(* Tests FB_Span.cloneTo, which processors use to keep a span that must outlive the original.
   A running span's context is taken through FB_Tracer.getSpanContext, tested in FB_TestTracer. *)
FUNCTION_BLOCK FB_TestSpan EXTENDS FB_TestSuite

THIS^.testCloneToCopiesEveryMember();
THIS^.testCloneToRejectsAssignedDestination();

(* cloneTo gives the copy its own copy of every member, so it outlives the source. *)
METHOD testCloneToCopiesEveryMember : REFERENCE TO FB_Test
VAR
	resource: FB_Resource('');
	idGenerator: FB_MockIdGenerator;
	provider: FB_TracerProvider_ForInspection(resource:=resource, idGenerator:=idGenerator, sampler:=TcOtlp_GVL.defaultSampler);
	scope: FB_InstrumentationScope('tracer.test', '1.0.0', '');
	tracer: FB_Tracer(scope:=scope, provider:=provider);
	pParent: POINTER TO FB_Span;
	pContext: POINTER TO FB_SpanContext;
	pSpan: POINTER TO FB_Span;
	pClone: POINTER TO FB_Span;
	pLink: POINTER TO FB_Link;
	pSourceLink: POINTER TO FB_Link;
	reason: E_SpanCloneFailureReason;
END_VAR
TcUnit.TEST('testCloneToCopiesEveryMember');
	IF resource.attributes.count = 0 THEN
		resource.attributes.setStringAttribute('host.id', 'PLC1');
	END_IF
	tracer.startSpan(name:='parent').build(pDest:=pParent);
	IF pParent <> 0 THEN tracer.getSpanContext(pSpan:=pParent, pDest:=pContext); END_IF
	tracer.startSpan(name:='work', kind:=E_SpanKind.SPAN_KIND_SERVER)
		.setParentUsingContext(pContext:=pContext)
		.addLink(pContext:=pContext)
		.setStringAttribute(key:='k', value:='v')
		.build(pDest:=pSpan);
	THIS^.AssertTrue(pSpan <> 0, 'Expected the span to build');
	IF pSpan <> 0 THEN
		// no builder sets timestamps; fixed values make the copy checkable
		pSpan^.startTimestamp := 1000;
		pSpan^.endTimestamp := 1500;
		tracer.setSpanStatusError(pSpan:=pSpan, message:='boom');
		pSpan^.links.reset();
		pSourceLink := pSpan^.links.next();

		THIS^.AssertTrue(pSpan^.cloneTo(pDest:=pClone, failureReason=>reason), 'Expected cloneTo to succeed');
		THIS^.AssertEquals_UDINT(TO_UDINT(E_SpanCloneFailureReason.NA), TO_UDINT(reason), 'Expected no failure');
		IF pClone <> 0 THEN
			THIS^.AssertTrue(pClone^.name <> 0 AND_THEN pClone^.name <> pSpan^.name, 'Expected a copied name');
			THIS^.AssertTrue(pClone^.traceId <> 0 AND_THEN pClone^.traceId <> pSpan^.traceId
				AND_THEN MEMCMP(ADR(pClone^.traceId^.bytes), ADR(pSpan^.traceId^.bytes), SIZEOF(pSpan^.traceId^.bytes)) = 0,
				'Expected a copied trace id');
			THIS^.AssertTrue(pClone^.spanId <> 0 AND_THEN pClone^.spanId <> pSpan^.spanId
				AND_THEN MEMCMP(ADR(pClone^.spanId^.bytes), ADR(pSpan^.spanId^.bytes), SIZEOF(pSpan^.spanId^.bytes)) = 0,
				'Expected a copied span id');
			THIS^.AssertTrue(pClone^.parentSpanId <> 0 AND_THEN pClone^.parentSpanId <> pSpan^.parentSpanId
				AND_THEN MEMCMP(ADR(pClone^.parentSpanId^.bytes), ADR(pSpan^.parentSpanId^.bytes), SIZEOF(pSpan^.parentSpanId^.bytes)) = 0,
				'Expected a copied parent span id');
			THIS^.AssertEquals_UDINT(TO_UDINT(E_SpanKind.SPAN_KIND_SERVER), TO_UDINT(pClone^.kind), 'Expected the kind');
			THIS^.AssertTrue(pClone^.startTimestamp = 1000 AND pClone^.endTimestamp = 1500, 'Expected the timestamps');
			THIS^.AssertEquals_UDINT(pSpan^.flags, pClone^.flags, 'Expected the flags');
			THIS^.AssertTrue(pClone^.status <> 0 AND_THEN pClone^.status <> pSpan^.status
				AND_THEN pClone^.status^.code = E_StatusCode.STATUS_CODE_ERROR
				AND_THEN pClone^.status^.message <> 0
				AND_THEN pClone^.status^.message <> pSpan^.status^.message,
				'Expected a copied error status');
			THIS^.AssertEquals_UDINT(pSpan^.attributes.count, pClone^.attributes.count, 'Expected the attributes');
			THIS^.AssertEquals_UDINT(1, pClone^.attributes.count, 'Expected one attribute');
			THIS^.AssertEquals_UDINT(1, pClone^.links.count, 'Expected one link');
			pClone^.links.reset();
			pLink := pClone^.links.next();
			THIS^.AssertTrue(pLink <> 0 AND_THEN pLink <> pSourceLink AND_THEN pLink^.spanId <> 0
				AND_THEN MEMCMP(ADR(pLink^.spanId^.bytes), ADR(pSourceLink^.spanId^.bytes), SIZEOF(pLink^.spanId^.bytes)) = 0,
				'Expected a copied link');
			THIS^.AssertEquals_UDINT(pSpan^.resource.attributes.count, pClone^.resource.attributes.count, 'Expected the resource');
			THIS^.AssertTrue(pClone^.resource.attributes.count > 0, 'Expected resource attributes to be copied');

			// the copy must stay valid once the source is gone
			pSpan^.delete(pSelf:=pSpan);
			THIS^.AssertEquals_STRING('work', pClone^.name^.pString^, 'Expected the name to outlive the source');
			THIS^.AssertEquals_STRING('boom', pClone^.status^.message^.pString^, 'Expected the message to outlive the source');
			pClone^.delete(pSelf:=pClone);
		END_IF
		IF pSpan <> 0 THEN pSpan^.delete(pSelf:=pSpan); END_IF
	END_IF
	IF pContext <> 0 THEN pContext^.delete(pSelf:=pContext); END_IF
	IF pParent <> 0 THEN pParent^.delete(pSelf:=pParent); END_IF
TcUnit.TEST_FINISHED();
END_METHOD

(* cloneTo refuses a destination that already holds a span and leaves it alone. *)
METHOD testCloneToRejectsAssignedDestination : REFERENCE TO FB_Test
VAR
	pSpan: POINTER TO FB_Span;
	pDest: POINTER TO FB_Span;
	reason: E_SpanCloneFailureReason;
END_VAR
TcUnit.TEST('testCloneToRejectsAssignedDestination');
	pSpan := __NEW(FB_Span);  // identity is irrelevant: only the destination check runs
	pDest := pSpan;  // deliberately assigned, so cloneTo must refuse it
	IF pSpan <> 0 THEN
		THIS^.AssertFalse(pSpan^.cloneTo(pDest:=pDest, failureReason=>reason), 'Expected cloneTo to fail');
		THIS^.AssertEquals_UDINT(
			TO_UDINT(E_SpanCloneFailureReason.DESTINATION_ALREADY_ASSIGNED),
			TO_UDINT(reason),
			'Expected DESTINATION_ALREADY_ASSIGNED'
		);
		THIS^.AssertTrue(pDest = pSpan, 'Expected the destination to be left alone');
		pSpan^.delete(pSelf:=pSpan);
	END_IF
TcUnit.TEST_FINISHED();
END_METHOD

END_FUNCTION_BLOCK

(* stored: Version 1.1.0.1
   POU FB_TestSpan: Id {db2f10cc-3e6d-4621-b34d-b5ee61137998}, SpecialFunc None
   Method testCloneToCopiesEveryMember: Id {4490e7af-97e3-416a-8e55-ef9dd747b048}
   Method testCloneToRejectsAssignedDestination: Id {ad9ae434-2120-4175-ad8f-7b344b3e8934} *)
